(* IEC 61131-3 sources: repolevel_ST_code_completion/dataset/project_code/Robotics_DynamicModel/TorqueLimitationDemo, 2 files *)

(* ---- AxisLimits.st ---- *)
TYPE AxisLimits :
STRUCT
	maxVelocity : LREAL;
	maxAcceleration : LREAL;
	maxDeceleration : LREAL;
	maxJerk : LREAL;
	maxTorque : LREAL;
END_STRUCT
END_TYPE

(* ---- TorqueLimitationDemoStates.st ---- *)
{attribute 'strict'}
TYPE TorqueLimitationDemoStates :
(
	PowerAxisGroup,
	InitializeDynamicModel,
	InitializeTestMovement,
	InitializeUnlimitedTorqueMovement,
	ExecuteUnlimitedTorqueMovement,
	InitializeLimitedTorqueMovement,
	ExecuteLimitedTorqueMovement,
	InitializeMovementWithLoad,
	ExecuteMovementWithLoad,
	FinalizeTestMovement,
	DemoFinished
);
END_TYPE
